(* CODESYS project Message.xml

Project tree, tasks and I/O mapping:
  visualisation Message
*)

// /Message
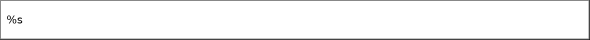
VISUALIZATION Message  // 590x40
VAR_IN_OUT
	scMessage 	: SC_LogMessage;
END_VAR
    Rectangle (0,0 590x40), "%s", text variable: scMessage.sMessage, colour toggle: scMessage.xError
END_VISUALIZATION
